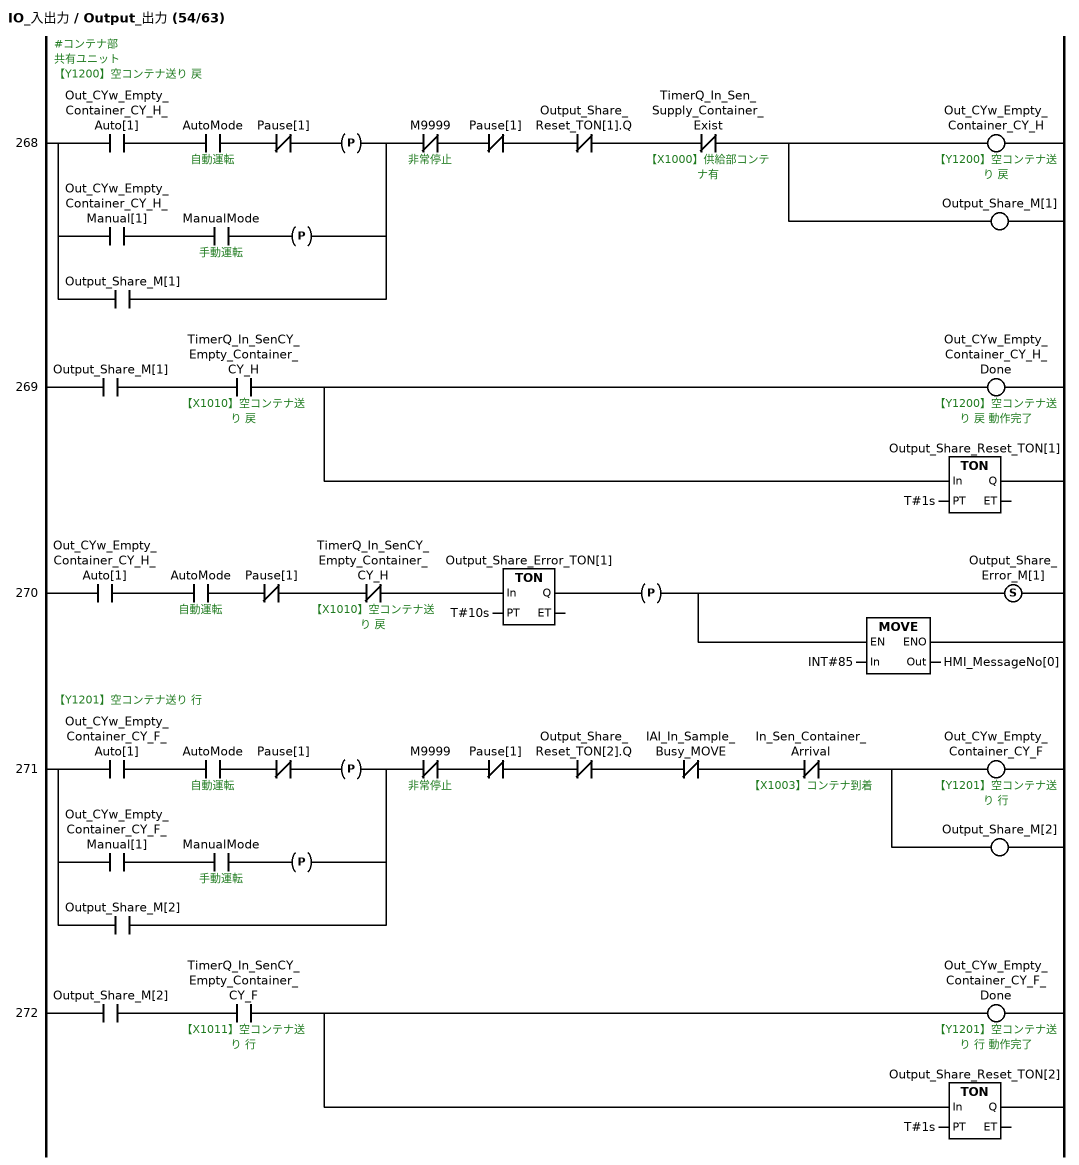
(* [picture p122: IO_入出力 / Output_出力, rungs 268-272] *)
(* Rung 268: #コンテナ部 / 共有ユニット / 【Y1200】空コンテナ送り 戻 *)
_e399(CLK := Out_CYw_Empty_Container_CY_H_Auto[1] AND AutoMode AND NOT Pause[1]);
_e400(CLK := Out_CYw_Empty_Container_CY_H_Manual[1] AND ManualMode);
_p401 := (_e399.Q OR _e400.Q OR Output_Share_M[1]) AND NOT M9999 AND NOT Pause[1] AND NOT Output_Share_Reset_TON[1].Q AND NOT TimerQ_In_Sen_Supply_Container_Exist;
Out_CYw_Empty_Container_CY_H := _p401;
Output_Share_M[1] := _p401;
(* Rung 269 *)
_p402 := Output_Share_M[1] AND TimerQ_In_SenCY_Empty_Container_CY_H;
Out_CYw_Empty_Container_CY_H_Done := _p402;
Output_Share_Reset_TON[1](In := _p402, PT := T#1s);
(* Rung 270 *)
Output_Share_Error_TON[1](In := Out_CYw_Empty_Container_CY_H_Auto[1] AND AutoMode AND NOT Pause[1] AND NOT TimerQ_In_SenCY_Empty_Container_CY_H, PT := T#10s);
_e403(CLK := Output_Share_Error_TON[1].Q);
IF _e403.Q THEN
    Output_Share_Error_M[1] := TRUE;
    HMI_MessageNo[0] := INT#85;
END_IF;
(* Rung 271: 【Y1201】空コンテナ送り 行 *)
_e404(CLK := Out_CYw_Empty_Container_CY_F_Auto[1] AND AutoMode AND NOT Pause[1]);
_e405(CLK := Out_CYw_Empty_Container_CY_F_Manual[1] AND ManualMode);
_p406 := (_e404.Q OR _e405.Q OR Output_Share_M[2]) AND NOT M9999 AND NOT Pause[1] AND NOT Output_Share_Reset_TON[2].Q AND NOT IAI_In_Sample_Busy_MOVE AND NOT In_Sen_Container_Arrival;
Out_CYw_Empty_Container_CY_F := _p406;
Output_Share_M[2] := _p406;
(* Rung 272 *)
_p407 := Output_Share_M[2] AND TimerQ_In_SenCY_Empty_Container_CY_F;
Out_CYw_Empty_Container_CY_F_Done := _p407;
Output_Share_Reset_TON[2](In := _p407, PT := T#1s);

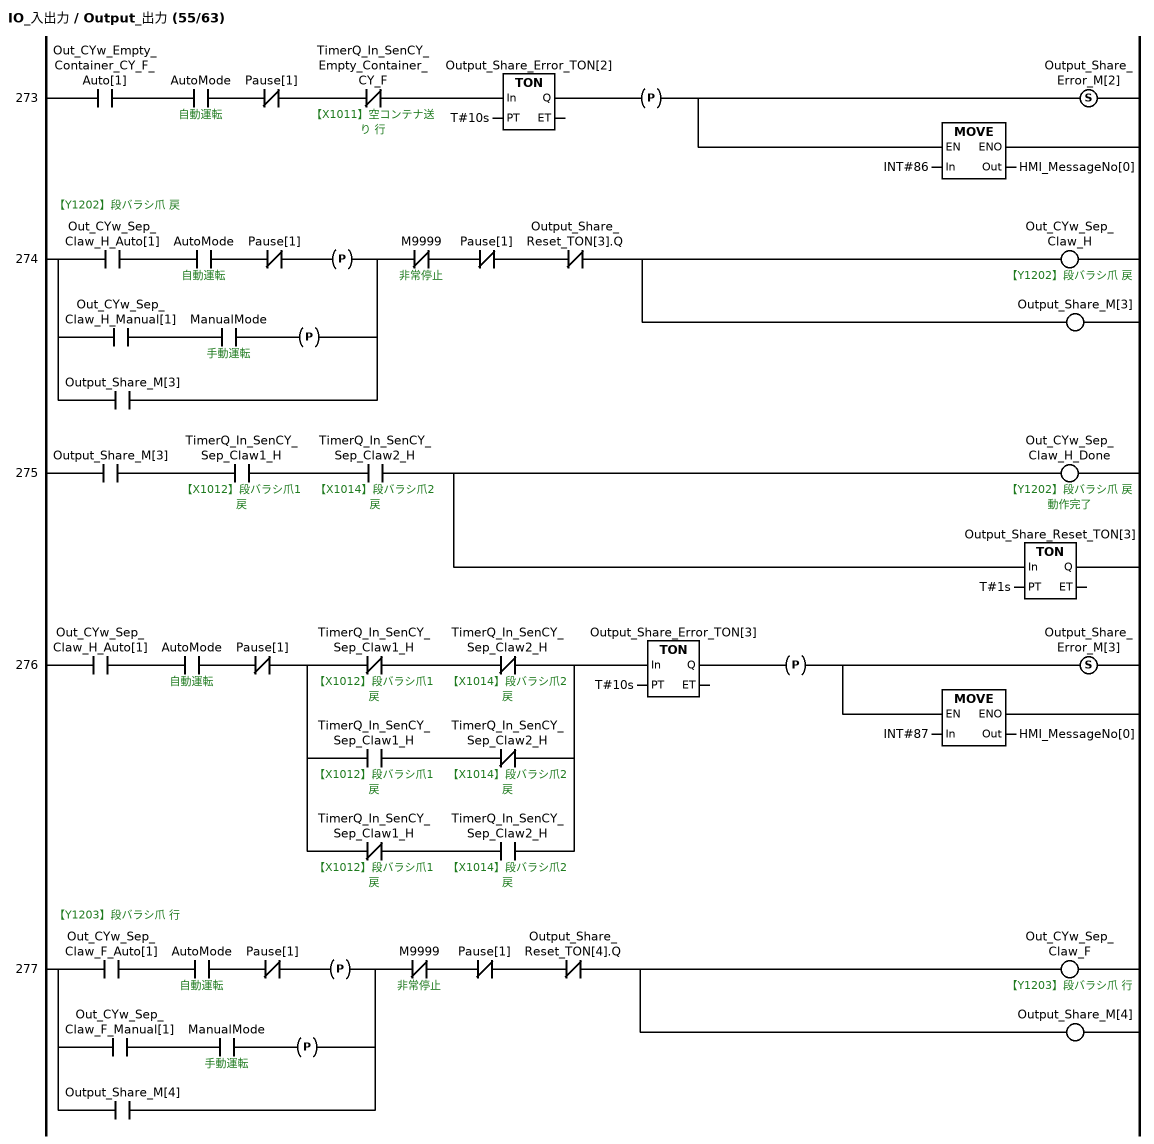
(* Rung 273 *)
Output_Share_Error_TON[2](In := Out_CYw_Empty_Container_CY_F_Auto[1] AND AutoMode AND NOT Pause[1] AND NOT TimerQ_In_SenCY_Empty_Container_CY_F, PT := T#10s);
_e408(CLK := Output_Share_Error_TON[2].Q);
IF _e408.Q THEN
    Output_Share_Error_M[2] := TRUE;
    HMI_MessageNo[0] := INT#86;
END_IF;
(* Rung 274: 【Y1202】段バラシ爪 戻 *)
_e409(CLK := Out_CYw_Sep_Claw_H_Auto[1] AND AutoMode AND NOT Pause[1]);
_e410(CLK := Out_CYw_Sep_Claw_H_Manual[1] AND ManualMode);
_p411 := (_e409.Q OR _e410.Q OR Output_Share_M[3]) AND NOT M9999 AND NOT Pause[1] AND NOT Output_Share_Reset_TON[3].Q;
Out_CYw_Sep_Claw_H := _p411;
Output_Share_M[3] := _p411;
(* Rung 275 *)
_p412 := Output_Share_M[3] AND TimerQ_In_SenCY_Sep_Claw1_H AND TimerQ_In_SenCY_Sep_Claw2_H;
Out_CYw_Sep_Claw_H_Done := _p412;
Output_Share_Reset_TON[3](In := _p412, PT := T#1s);
(* Rung 276 *)
Output_Share_Error_TON[3](In := Out_CYw_Sep_Claw_H_Auto[1] AND AutoMode AND NOT Pause[1] AND ((NOT TimerQ_In_SenCY_Sep_Claw1_H AND NOT TimerQ_In_SenCY_Sep_Claw2_H) OR (TimerQ_In_SenCY_Sep_Claw1_H AND NOT TimerQ_In_SenCY_Sep_Claw2_H) OR (NOT TimerQ_In_SenCY_Sep_Claw1_H AND TimerQ_In_SenCY_Sep_Claw2_H)), PT := T#10s);
_e413(CLK := Output_Share_Error_TON[3].Q);
IF _e413.Q THEN
    Output_Share_Error_M[3] := TRUE;
    HMI_MessageNo[0] := INT#87;
END_IF;
(* Rung 277: 【Y1203】段バラシ爪 行 *)
_e414(CLK := Out_CYw_Sep_Claw_F_Auto[1] AND AutoMode AND NOT Pause[1]);
_e415(CLK := Out_CYw_Sep_Claw_F_Manual[1] AND ManualMode);
_p416 := (_e414.Q OR _e415.Q OR Output_Share_M[4]) AND NOT M9999 AND NOT Pause[1] AND NOT Output_Share_Reset_TON[4].Q;
Out_CYw_Sep_Claw_F := _p416;
Output_Share_M[4] := _p416;

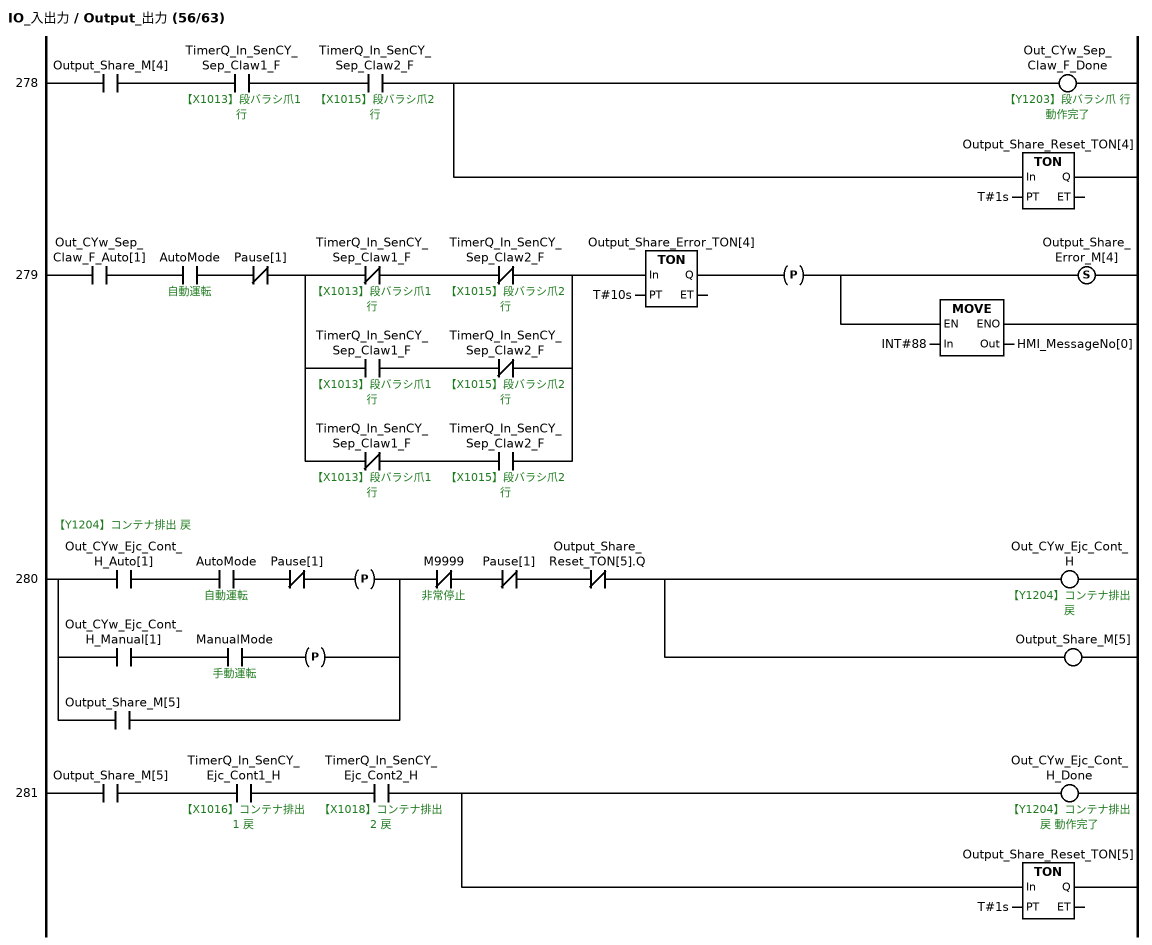
(* Rung 278 *)
_p417 := Output_Share_M[4] AND TimerQ_In_SenCY_Sep_Claw1_F AND TimerQ_In_SenCY_Sep_Claw2_F;
Out_CYw_Sep_Claw_F_Done := _p417;
Output_Share_Reset_TON[4](In := _p417, PT := T#1s);
(* Rung 279 *)
Output_Share_Error_TON[4](In := Out_CYw_Sep_Claw_F_Auto[1] AND AutoMode AND NOT Pause[1] AND ((NOT TimerQ_In_SenCY_Sep_Claw1_F AND NOT TimerQ_In_SenCY_Sep_Claw2_F) OR (TimerQ_In_SenCY_Sep_Claw1_F AND NOT TimerQ_In_SenCY_Sep_Claw2_F) OR (NOT TimerQ_In_SenCY_Sep_Claw1_F AND TimerQ_In_SenCY_Sep_Claw2_F)), PT := T#10s);
_e418(CLK := Output_Share_Error_TON[4].Q);
IF _e418.Q THEN
    Output_Share_Error_M[4] := TRUE;
    HMI_MessageNo[0] := INT#88;
END_IF;
(* Rung 280: 【Y1204】コンテナ排出 戻 *)
_e419(CLK := Out_CYw_Ejc_Cont_H_Auto[1] AND AutoMode AND NOT Pause[1]);
_e420(CLK := Out_CYw_Ejc_Cont_H_Manual[1] AND ManualMode);
_p421 := (_e419.Q OR _e420.Q OR Output_Share_M[5]) AND NOT M9999 AND NOT Pause[1] AND NOT Output_Share_Reset_TON[5].Q;
Out_CYw_Ejc_Cont_H := _p421;
Output_Share_M[5] := _p421;
(* Rung 281 *)
_p422 := Output_Share_M[5] AND TimerQ_In_SenCY_Ejc_Cont1_H AND TimerQ_In_SenCY_Ejc_Cont2_H;
Out_CYw_Ejc_Cont_H_Done := _p422;
Output_Share_Reset_TON[5](In := _p422, PT := T#1s);

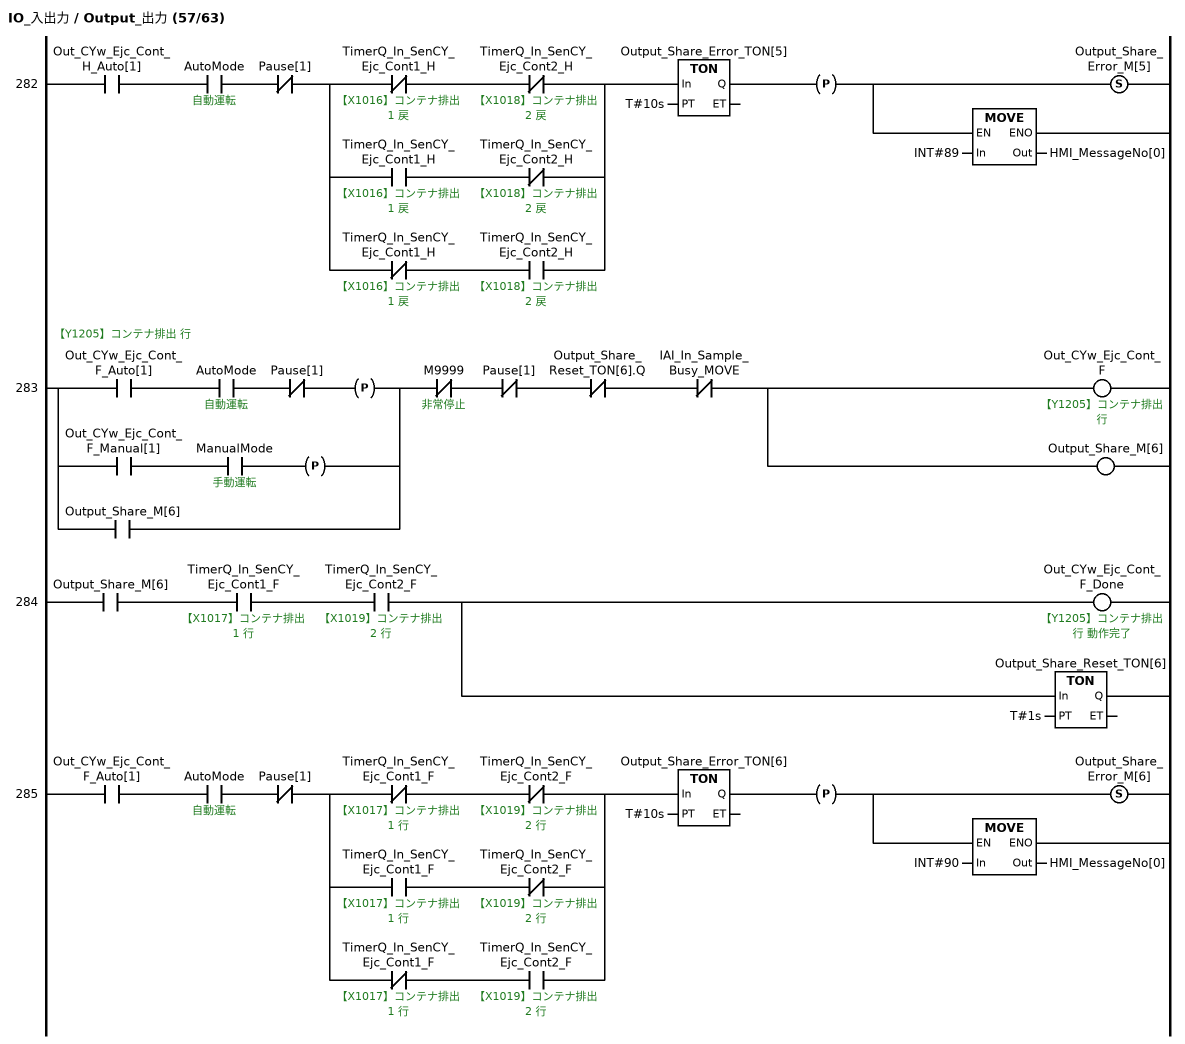
(* Rung 282 *)
Output_Share_Error_TON[5](In := Out_CYw_Ejc_Cont_H_Auto[1] AND AutoMode AND NOT Pause[1] AND ((NOT TimerQ_In_SenCY_Ejc_Cont1_H AND NOT TimerQ_In_SenCY_Ejc_Cont2_H) OR (TimerQ_In_SenCY_Ejc_Cont1_H AND NOT TimerQ_In_SenCY_Ejc_Cont2_H) OR (NOT TimerQ_In_SenCY_Ejc_Cont1_H AND TimerQ_In_SenCY_Ejc_Cont2_H)), PT := T#10s);
_e423(CLK := Output_Share_Error_TON[5].Q);
IF _e423.Q THEN
    Output_Share_Error_M[5] := TRUE;
    HMI_MessageNo[0] := INT#89;
END_IF;
(* Rung 283: 【Y1205】コンテナ排出 行 *)
_e424(CLK := Out_CYw_Ejc_Cont_F_Auto[1] AND AutoMode AND NOT Pause[1]);
_e425(CLK := Out_CYw_Ejc_Cont_F_Manual[1] AND ManualMode);
_p426 := (_e424.Q OR _e425.Q OR Output_Share_M[6]) AND NOT M9999 AND NOT Pause[1] AND NOT Output_Share_Reset_TON[6].Q AND NOT IAI_In_Sample_Busy_MOVE;
Out_CYw_Ejc_Cont_F := _p426;
Output_Share_M[6] := _p426;
(* Rung 284 *)
_p427 := Output_Share_M[6] AND TimerQ_In_SenCY_Ejc_Cont1_F AND TimerQ_In_SenCY_Ejc_Cont2_F;
Out_CYw_Ejc_Cont_F_Done := _p427;
Output_Share_Reset_TON[6](In := _p427, PT := T#1s);
(* Rung 285 *)
Output_Share_Error_TON[6](In := Out_CYw_Ejc_Cont_F_Auto[1] AND AutoMode AND NOT Pause[1] AND ((NOT TimerQ_In_SenCY_Ejc_Cont1_F AND NOT TimerQ_In_SenCY_Ejc_Cont2_F) OR (TimerQ_In_SenCY_Ejc_Cont1_F AND NOT TimerQ_In_SenCY_Ejc_Cont2_F) OR (NOT TimerQ_In_SenCY_Ejc_Cont1_F AND TimerQ_In_SenCY_Ejc_Cont2_F)), PT := T#10s);
_e428(CLK := Output_Share_Error_TON[6].Q);
IF _e428.Q THEN
    Output_Share_Error_M[6] := TRUE;
    HMI_MessageNo[0] := INT#90;
END_IF;

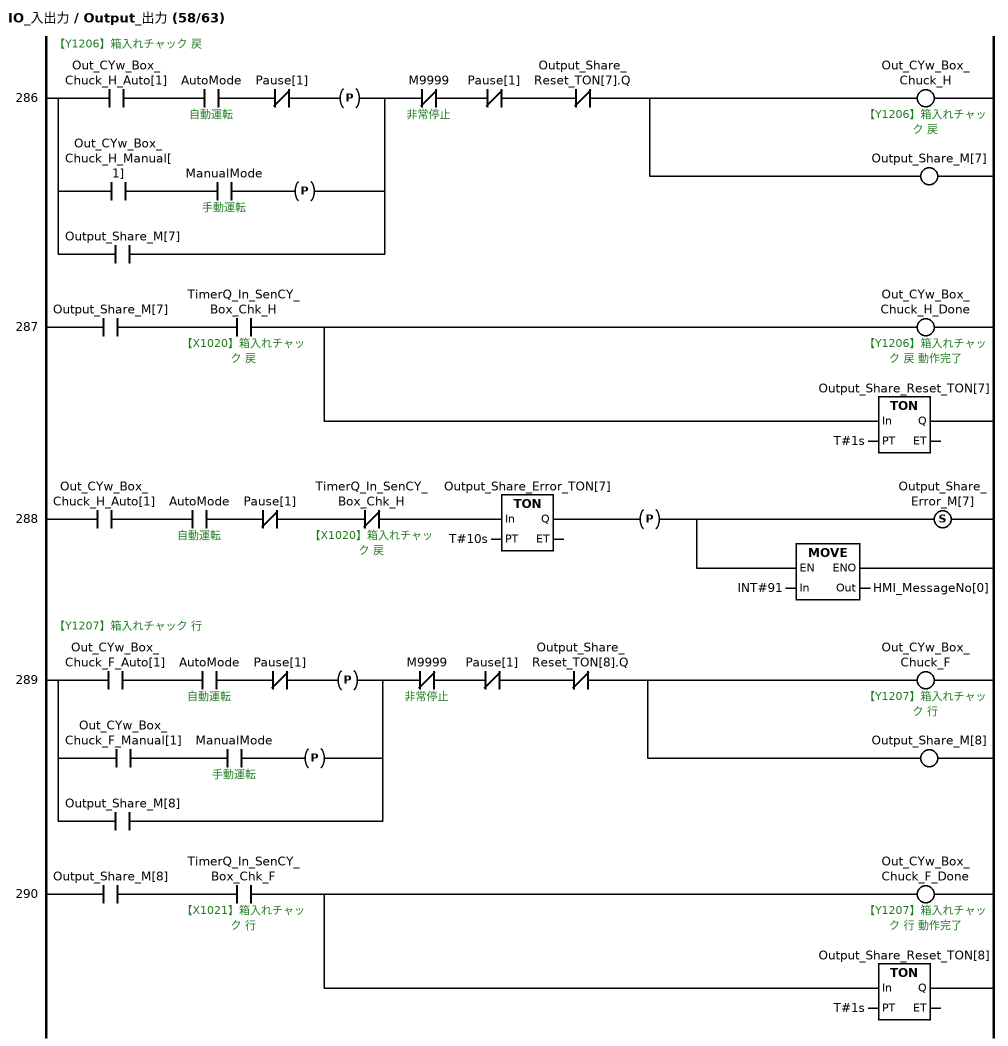
(* Rung 286: 【Y1206】箱入れチャック 戻 *)
_e429(CLK := Out_CYw_Box_Chuck_H_Auto[1] AND AutoMode AND NOT Pause[1]);
_e430(CLK := Out_CYw_Box_Chuck_H_Manual[1] AND ManualMode);
_p431 := (_e429.Q OR _e430.Q OR Output_Share_M[7]) AND NOT M9999 AND NOT Pause[1] AND NOT Output_Share_Reset_TON[7].Q;
Out_CYw_Box_Chuck_H := _p431;
Output_Share_M[7] := _p431;
(* Rung 287 *)
Out_CYw_Box_Chuck_H_Done := Output_Share_M[7] AND TimerQ_In_SenCY_Box_Chk_H;
Output_Share_Reset_TON[7](In := Output_Share_M[7] AND TimerQ_In_SenCY_Box_Chk_H, PT := T#1s);
(* Rung 288 *)
Output_Share_Error_TON[7](In := Out_CYw_Box_Chuck_H_Auto[1] AND AutoMode AND NOT Pause[1] AND NOT TimerQ_In_SenCY_Box_Chk_H, PT := T#10s);
_e432(CLK := Output_Share_Error_TON[7].Q);
IF _e432.Q THEN
    Output_Share_Error_M[7] := TRUE;
    HMI_MessageNo[0] := INT#91;
END_IF;
(* Rung 289: 【Y1207】箱入れチャック 行 *)
_e433(CLK := Out_CYw_Box_Chuck_F_Auto[1] AND AutoMode AND NOT Pause[1]);
_e434(CLK := Out_CYw_Box_Chuck_F_Manual[1] AND ManualMode);
_p435 := (_e433.Q OR _e434.Q OR Output_Share_M[8]) AND NOT M9999 AND NOT Pause[1] AND NOT Output_Share_Reset_TON[8].Q;
Out_CYw_Box_Chuck_F := _p435;
Output_Share_M[8] := _p435;
(* Rung 290 *)
Out_CYw_Box_Chuck_F_Done := Output_Share_M[8] AND TimerQ_In_SenCY_Box_Chk_F;
Output_Share_Reset_TON[8](In := Output_Share_M[8] AND TimerQ_In_SenCY_Box_Chk_F, PT := T#1s);

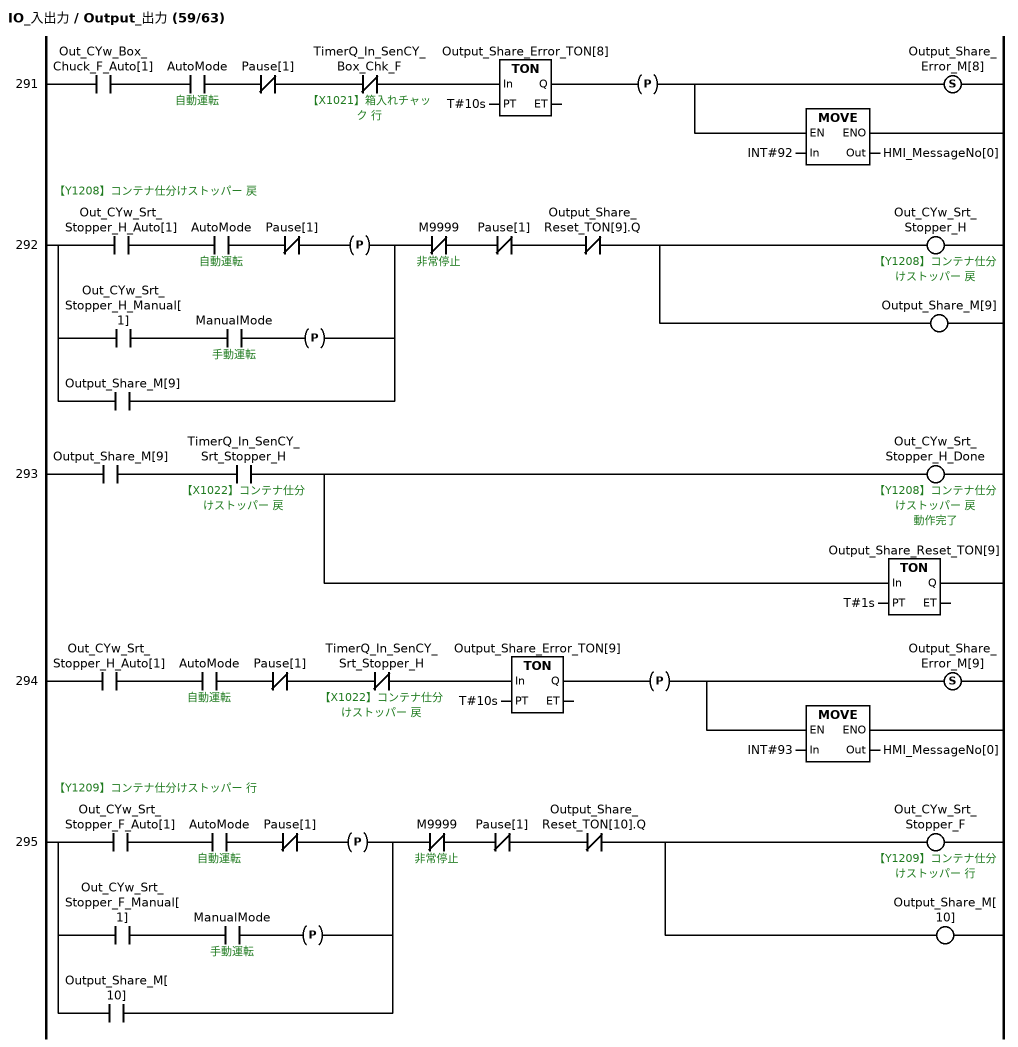
(* Rung 291 *)
Output_Share_Error_TON[8](In := Out_CYw_Box_Chuck_F_Auto[1] AND AutoMode AND NOT Pause[1] AND NOT TimerQ_In_SenCY_Box_Chk_F, PT := T#10s);
_e436(CLK := Output_Share_Error_TON[8].Q);
IF _e436.Q THEN
    Output_Share_Error_M[8] := TRUE;
    HMI_MessageNo[0] := INT#92;
END_IF;
(* Rung 292: 【Y1208】コンテナ仕分けストッパー 戻 *)
_e437(CLK := Out_CYw_Srt_Stopper_H_Auto[1] AND AutoMode AND NOT Pause[1]);
_e438(CLK := Out_CYw_Srt_Stopper_H_Manual[1] AND ManualMode);
_p439 := (_e437.Q OR _e438.Q OR Output_Share_M[9]) AND NOT M9999 AND NOT Pause[1] AND NOT Output_Share_Reset_TON[9].Q;
Out_CYw_Srt_Stopper_H := _p439;
Output_Share_M[9] := _p439;
(* Rung 293 *)
_p440 := Output_Share_M[9] AND TimerQ_In_SenCY_Srt_Stopper_H;
Out_CYw_Srt_Stopper_H_Done := _p440;
Output_Share_Reset_TON[9](In := _p440, PT := T#1s);
(* Rung 294 *)
Output_Share_Error_TON[9](In := Out_CYw_Srt_Stopper_H_Auto[1] AND AutoMode AND NOT Pause[1] AND NOT TimerQ_In_SenCY_Srt_Stopper_H, PT := T#10s);
_e441(CLK := Output_Share_Error_TON[9].Q);
IF _e441.Q THEN
    Output_Share_Error_M[9] := TRUE;
    HMI_MessageNo[0] := INT#93;
END_IF;
(* Rung 295: 【Y1209】コンテナ仕分けストッパー 行 *)
_e442(CLK := Out_CYw_Srt_Stopper_F_Auto[1] AND AutoMode AND NOT Pause[1]);
_e443(CLK := Out_CYw_Srt_Stopper_F_Manual[1] AND ManualMode);
_p444 := (_e442.Q OR _e443.Q OR Output_Share_M[10]) AND NOT M9999 AND NOT Pause[1] AND NOT Output_Share_Reset_TON[10].Q;
Out_CYw_Srt_Stopper_F := _p444;
Output_Share_M[10] := _p444;

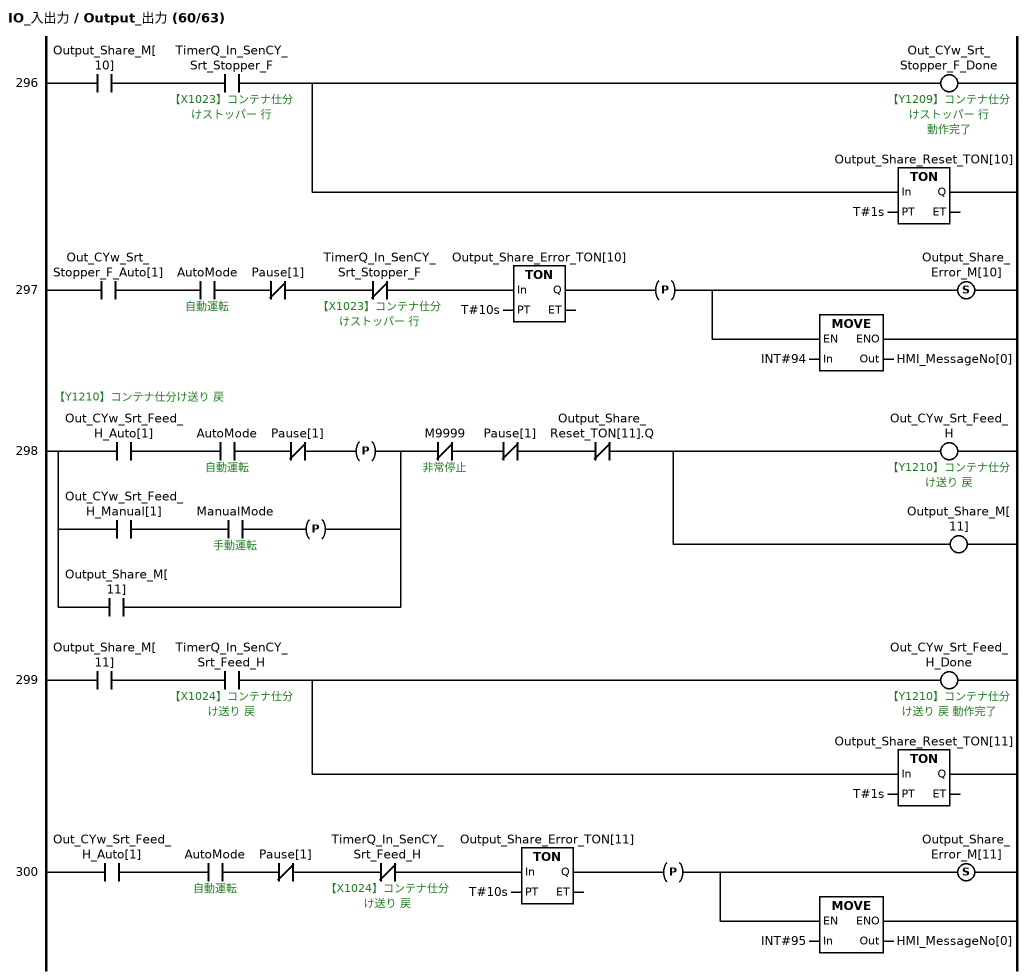
(* Rung 296 *)
_p445 := Output_Share_M[10] AND TimerQ_In_SenCY_Srt_Stopper_F;
Out_CYw_Srt_Stopper_F_Done := _p445;
Output_Share_Reset_TON[10](In := _p445, PT := T#1s);
(* Rung 297 *)
Output_Share_Error_TON[10](In := Out_CYw_Srt_Stopper_F_Auto[1] AND AutoMode AND NOT Pause[1] AND NOT TimerQ_In_SenCY_Srt_Stopper_F, PT := T#10s);
_e446(CLK := Output_Share_Error_TON[10].Q);
IF _e446.Q THEN
    Output_Share_Error_M[10] := TRUE;
    HMI_MessageNo[0] := INT#94;
END_IF;
(* Rung 298: 【Y1210】コンテナ仕分け送り 戻 *)
_e447(CLK := Out_CYw_Srt_Feed_H_Auto[1] AND AutoMode AND NOT Pause[1]);
_e448(CLK := Out_CYw_Srt_Feed_H_Manual[1] AND ManualMode);
_p449 := (_e447.Q OR _e448.Q OR Output_Share_M[11]) AND NOT M9999 AND NOT Pause[1] AND NOT Output_Share_Reset_TON[11].Q;
Out_CYw_Srt_Feed_H := _p449;
Output_Share_M[11] := _p449;
(* Rung 299 *)
_p450 := Output_Share_M[11] AND TimerQ_In_SenCY_Srt_Feed_H;
Out_CYw_Srt_Feed_H_Done := _p450;
Output_Share_Reset_TON[11](In := _p450, PT := T#1s);
(* Rung 300 *)
Output_Share_Error_TON[11](In := Out_CYw_Srt_Feed_H_Auto[1] AND AutoMode AND NOT Pause[1] AND NOT TimerQ_In_SenCY_Srt_Feed_H, PT := T#10s);
_e451(CLK := Output_Share_Error_TON[11].Q);
IF _e451.Q THEN
    Output_Share_Error_M[11] := TRUE;
    HMI_MessageNo[0] := INT#95;
END_IF;

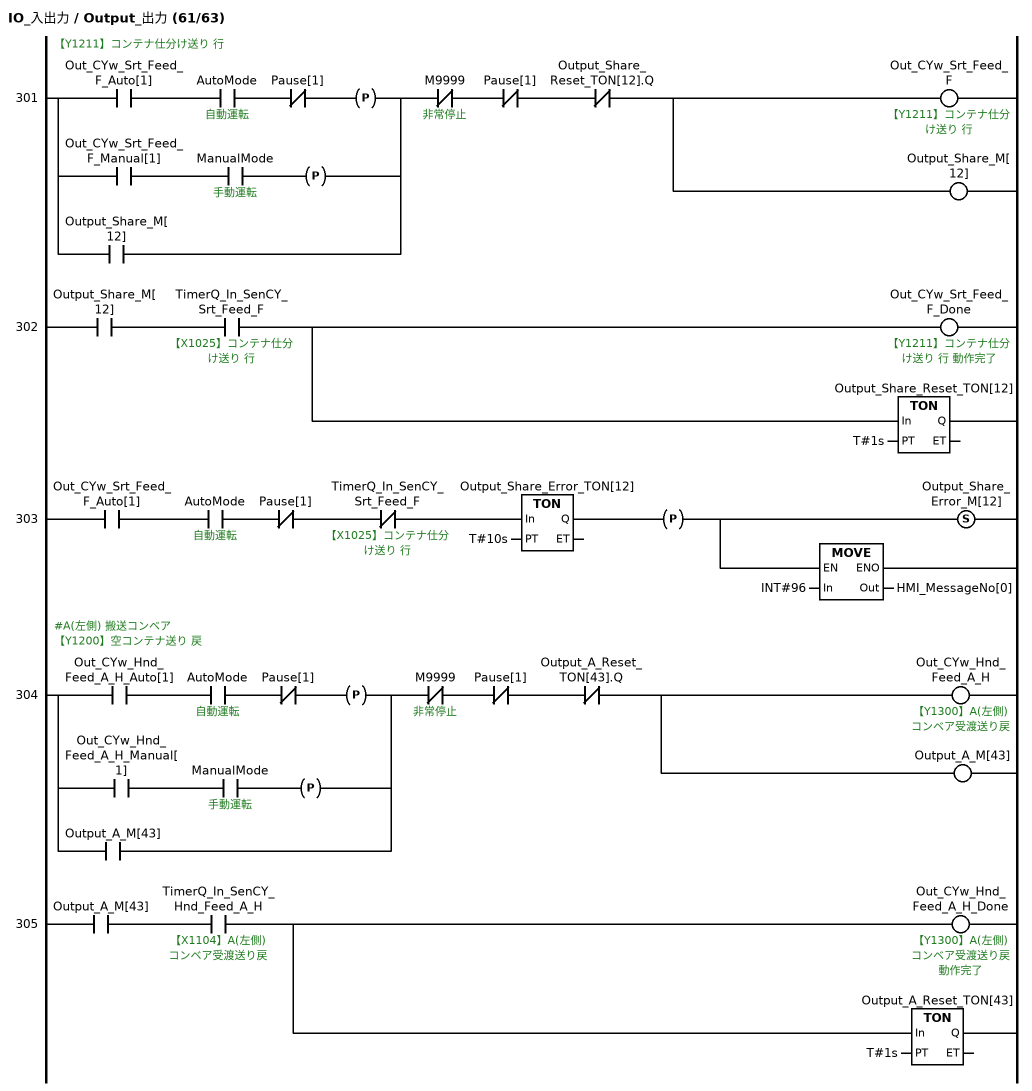
(* Rung 301: 【Y1211】コンテナ仕分け送り 行 *)
_e452(CLK := Out_CYw_Srt_Feed_F_Auto[1] AND AutoMode AND NOT Pause[1]);
_e453(CLK := Out_CYw_Srt_Feed_F_Manual[1] AND ManualMode);
_p454 := (_e452.Q OR _e453.Q OR Output_Share_M[12]) AND NOT M9999 AND NOT Pause[1] AND NOT Output_Share_Reset_TON[12].Q;
Out_CYw_Srt_Feed_F := _p454;
Output_Share_M[12] := _p454;
(* Rung 302 *)
_p455 := Output_Share_M[12] AND TimerQ_In_SenCY_Srt_Feed_F;
Out_CYw_Srt_Feed_F_Done := _p455;
Output_Share_Reset_TON[12](In := _p455, PT := T#1s);
(* Rung 303 *)
Output_Share_Error_TON[12](In := Out_CYw_Srt_Feed_F_Auto[1] AND AutoMode AND NOT Pause[1] AND NOT TimerQ_In_SenCY_Srt_Feed_F, PT := T#10s);
_e456(CLK := Output_Share_Error_TON[12].Q);
IF _e456.Q THEN
    Output_Share_Error_M[12] := TRUE;
    HMI_MessageNo[0] := INT#96;
END_IF;
(* Rung 304: #A(左側) 搬送コンベア / 【Y1200】空コンテナ送り 戻 *)
_e457(CLK := Out_CYw_Hnd_Feed_A_H_Auto[1] AND AutoMode AND NOT Pause[1]);
_e458(CLK := Out_CYw_Hnd_Feed_A_H_Manual[1] AND ManualMode);
_p459 := (_e457.Q OR _e458.Q OR Output_A_M[43]) AND NOT M9999 AND NOT Pause[1] AND NOT Output_A_Reset_TON[43].Q;
Out_CYw_Hnd_Feed_A_H := _p459;
Output_A_M[43] := _p459;
(* Rung 305 *)
Out_CYw_Hnd_Feed_A_H_Done := Output_A_M[43] AND TimerQ_In_SenCY_Hnd_Feed_A_H;
Output_A_Reset_TON[43](In := Output_A_M[43] AND TimerQ_In_SenCY_Hnd_Feed_A_H, PT := T#1s);

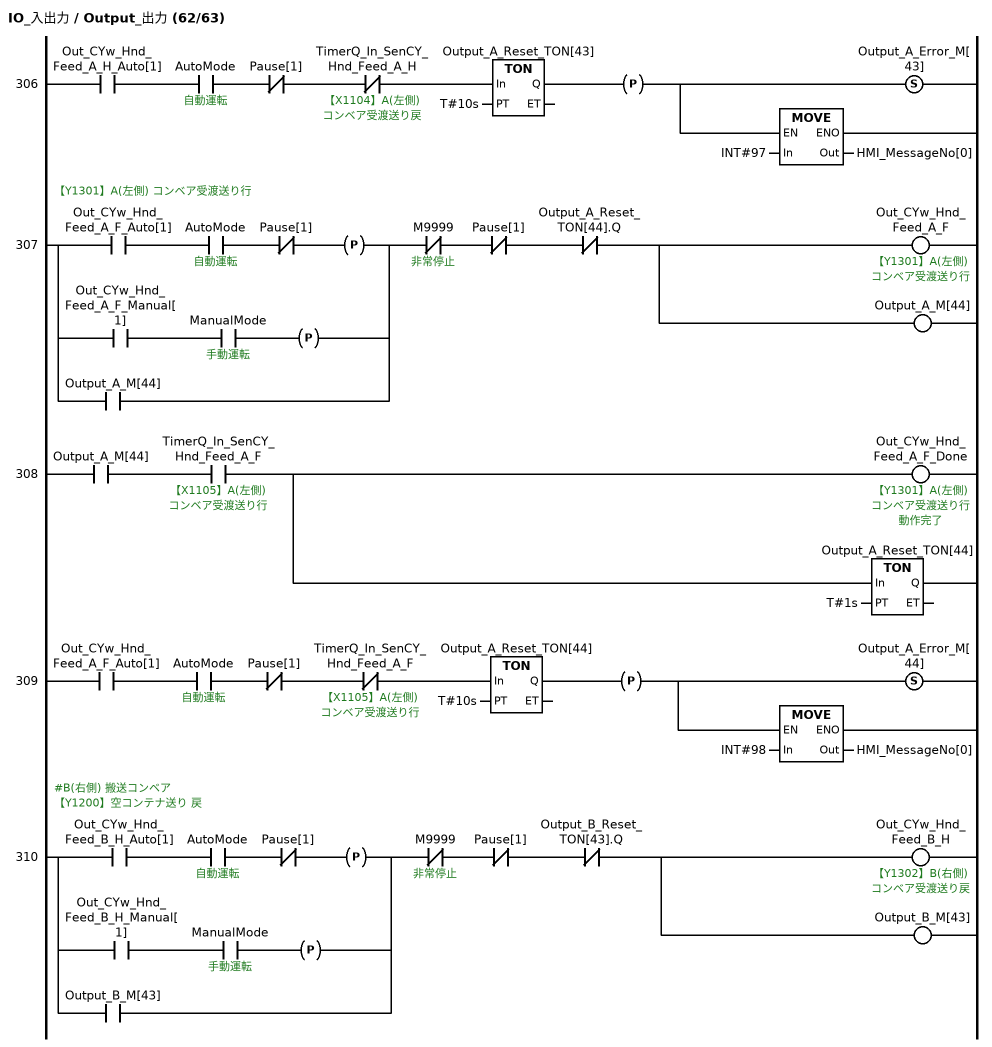
(* Rung 306 *)
Output_A_Reset_TON[43](In := Out_CYw_Hnd_Feed_A_H_Auto[1] AND AutoMode AND NOT Pause[1] AND NOT TimerQ_In_SenCY_Hnd_Feed_A_H, PT := T#10s);
_e460(CLK := Output_A_Reset_TON[43].Q);
IF _e460.Q THEN
    Output_A_Error_M[43] := TRUE;
    HMI_MessageNo[0] := INT#97;
END_IF;
(* Rung 307: 【Y1301】A(左側) コンベア受渡送り行 *)
_e461(CLK := Out_CYw_Hnd_Feed_A_F_Auto[1] AND AutoMode AND NOT Pause[1]);
_e462(CLK := Out_CYw_Hnd_Feed_A_F_Manual[1] AND ManualMode);
_p463 := (_e461.Q OR _e462.Q OR Output_A_M[44]) AND NOT M9999 AND NOT Pause[1] AND NOT Output_A_Reset_TON[44].Q;
Out_CYw_Hnd_Feed_A_F := _p463;
Output_A_M[44] := _p463;
(* Rung 308 *)
Out_CYw_Hnd_Feed_A_F_Done := Output_A_M[44] AND TimerQ_In_SenCY_Hnd_Feed_A_F;
Output_A_Reset_TON[44](In := Output_A_M[44] AND TimerQ_In_SenCY_Hnd_Feed_A_F, PT := T#1s);
(* Rung 309 *)
Output_A_Reset_TON[44](In := Out_CYw_Hnd_Feed_A_F_Auto[1] AND AutoMode AND NOT Pause[1] AND NOT TimerQ_In_SenCY_Hnd_Feed_A_F, PT := T#10s);
_e464(CLK := Output_A_Reset_TON[44].Q);
IF _e464.Q THEN
    Output_A_Error_M[44] := TRUE;
    HMI_MessageNo[0] := INT#98;
END_IF;
(* Rung 310: #B(右側) 搬送コンベア / 【Y1200】空コンテナ送り 戻 *)
_e465(CLK := Out_CYw_Hnd_Feed_B_H_Auto[1] AND AutoMode AND NOT Pause[1]);
_e466(CLK := Out_CYw_Hnd_Feed_B_H_Manual[1] AND ManualMode);
_p467 := (_e465.Q OR _e466.Q OR Output_B_M[43]) AND NOT M9999 AND NOT Pause[1] AND NOT Output_B_Reset_TON[43].Q;
Out_CYw_Hnd_Feed_B_H := _p467;
Output_B_M[43] := _p467;

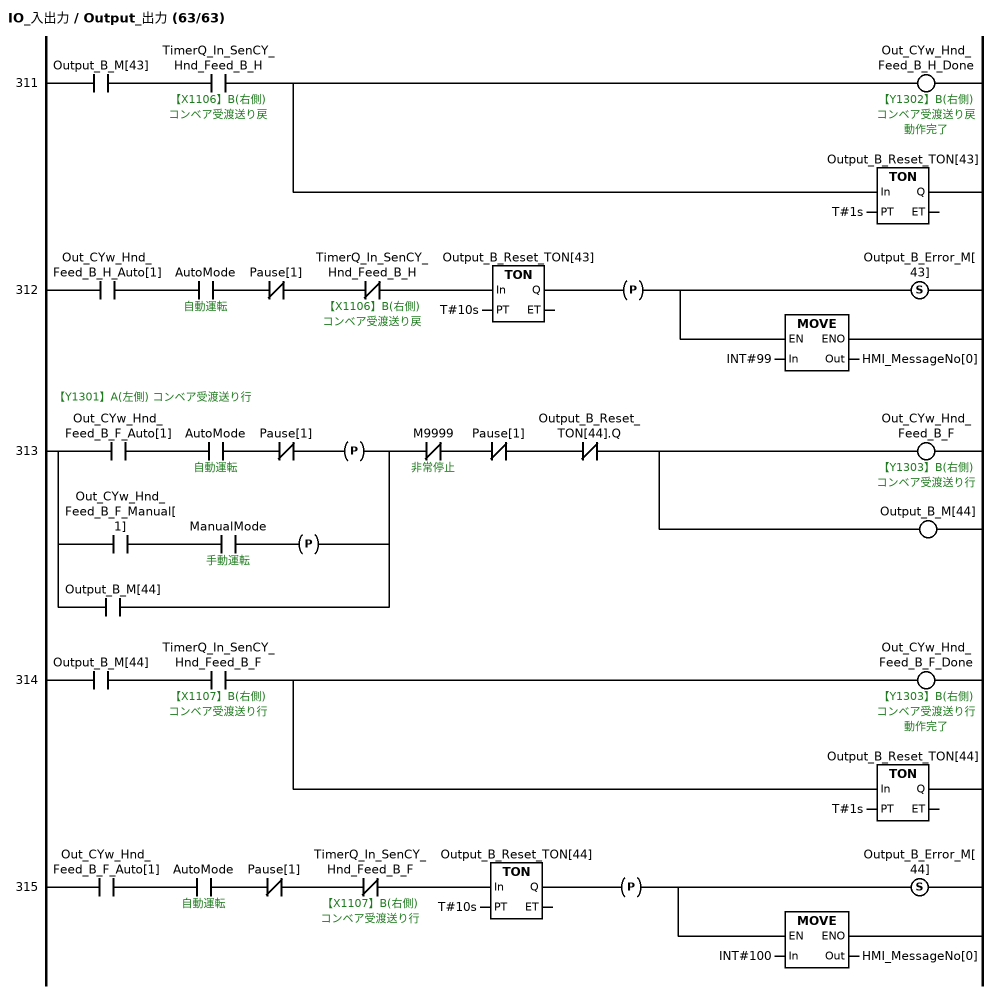
(* Rung 311 *)
Out_CYw_Hnd_Feed_B_H_Done := Output_B_M[43] AND TimerQ_In_SenCY_Hnd_Feed_B_H;
Output_B_Reset_TON[43](In := Output_B_M[43] AND TimerQ_In_SenCY_Hnd_Feed_B_H, PT := T#1s);
(* Rung 312 *)
Output_B_Reset_TON[43](In := Out_CYw_Hnd_Feed_B_H_Auto[1] AND AutoMode AND NOT Pause[1] AND NOT TimerQ_In_SenCY_Hnd_Feed_B_H, PT := T#10s);
_e468(CLK := Output_B_Reset_TON[43].Q);
IF _e468.Q THEN
    Output_B_Error_M[43] := TRUE;
    HMI_MessageNo[0] := INT#99;
END_IF;
(* Rung 313: 【Y1301】A(左側) コンベア受渡送り行 *)
_e469(CLK := Out_CYw_Hnd_Feed_B_F_Auto[1] AND AutoMode AND NOT Pause[1]);
_e470(CLK := Out_CYw_Hnd_Feed_B_F_Manual[1] AND ManualMode);
_p471 := (_e469.Q OR _e470.Q OR Output_B_M[44]) AND NOT M9999 AND NOT Pause[1] AND NOT Output_B_Reset_TON[44].Q;
Out_CYw_Hnd_Feed_B_F := _p471;
Output_B_M[44] := _p471;
(* Rung 314 *)
Out_CYw_Hnd_Feed_B_F_Done := Output_B_M[44] AND TimerQ_In_SenCY_Hnd_Feed_B_F;
Output_B_Reset_TON[44](In := Output_B_M[44] AND TimerQ_In_SenCY_Hnd_Feed_B_F, PT := T#1s);
(* Rung 315 *)
Output_B_Reset_TON[44](In := Out_CYw_Hnd_Feed_B_F_Auto[1] AND AutoMode AND NOT Pause[1] AND NOT TimerQ_In_SenCY_Hnd_Feed_B_F, PT := T#10s);
_e472(CLK := Output_B_Reset_TON[44].Q);
IF _e472.Q THEN
    Output_B_Error_M[44] := TRUE;
    HMI_MessageNo[0] := INT#100;
END_IF;
END_PROGRAM

# Device HMI_NA5_0 (NA): not converted